Staubli VAL3: _btnColor.pgx

public program _btnColor(num x_nSelType, string x_sHtml)
begin
  switch x_nSelType
    case 1
      userPageSet(x_sHtml,"btn7","style.backgroundColor","#7CB5FF")
      userPageSet(x_sHtml,"btn7","style.color","#FFFFFF")
      userPageSet(x_sHtml,"btn8","style.backgroundColor","#FFFFFF")
      userPageSet(x_sHtml,"btn8","style.color","#838A8F")
    break
    case 2
      userPageSet(x_sHtml,"btn8","style.backgroundColor","#7CB5FF")
      userPageSet(x_sHtml,"btn8","style.color","#FFFFFF")
      userPageSet(x_sHtml,"btn7","style.backgroundColor","#FFFFFF")
      userPageSet(x_sHtml,"btn7","style.color","#838A8F")
    break
  endSwitch

end
